SUBAPPLICATION SoftKeySR_PC_B_OPC_LOC (* Wie SoftKeySR_PC_B_OPC, aber Zustand lokal per PUBLISH (ein Geraet, Methoden per localhost) *)
  (* Standard: 61499-2; Description: Copyright (c) 2026 Meisterschulen am Ostbahnhof This program and the accompanying materials are made available under the terms of the Eclipse Public License 2.0 which is available at https://www.eclipse.org/legal/epl-2.0/ SPDX-License-Identifier: EPL-2.0 *)
  (* Version 1.3, 2026-11-25, Franz Höpfinger, Meisterschulen am Ostbahnhof, SERVER_0 -> MyLib::net::SERVER_0_QO (IND nur bei QO=TRUE, RSP intern). Ein gescheitertes RSP meldet IND mit QO=FALSE, direkt IND->RSP ergab eine Endlosschleife. *)
  (* Version 1.2, 2026-10-18, Franz Höpfinger, Meisterschulen am Ostbahnhof, Lokale Variante von SoftKeySR_PC_B_OPC: lokales PUBLISH statt Remote-WRITE (CLIENT) *)
  (* Version 1.1, 2026-09-09, Franz Höpfinger, Meisterschulen am Ostbahnhof, Fix: beide SERVER_0.RSP waren nie verdrahtet - blockierten je bis zu 4s den OPC-UA-Server-Thread (haelt open62541s globalen serviceMutex), verzoegerte dadurch JEDE OPC-UA-Statusmeldung projektweit. IND->RSP direkt verdrahtet. Siehe OPC_UA_VERNETZUNG.md Punkt 12. *)
  (* Version 1.0, 2026-09-03, Franz Höpfinger, Meisterschulen am Ostbahnhof, initial API and implementation and/or initial documentation *)
  PACKAGE MyLib::sys;
  IMPORT logiBUS::io::DQ::logiBUS_DO;
  IMPORT logiBUS::io::DQ::logiBUS_DO_S;
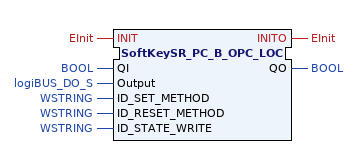
  EVENT_INPUT
    INIT : EInit; (* Initialization Request *)
  END_EVENT
  EVENT_OUTPUT
    INITO : EInit; (* Initialization Confirm *)
  END_EVENT
  VAR_INPUT
    QI : BOOL := TRUE; (* Quality Input - TRUE to enable service *)
    Output : logiBUS::io::DQ::logiBUS_DO_S := logiBUS_DO::Invalid; (* Identify the Output Output_Q1..Q8 *)
    ID_SET_METHOD : WSTRING; (* Lokale Methodenadresse (ACTION=CREATE_METHOD) fuer den Set-Methodenaufruf, wird von Geraet A per CALL_METHOD aufgerufen *)
    ID_RESET_METHOD : WSTRING; (* Lokale Methodenadresse (ACTION=CREATE_METHOD) fuer den Reset-Methodenaufruf, wird von Geraet A per CALL_METHOD aufgerufen *)
    ID_STATE_WRITE : WSTRING; (* Lokale Knotenadresse (BOOL, ACTION=WRITE) fuer den Zustand *)
  END_VAR
  VAR_OUTPUT
    QO : BOOL; (* Quality Output - TRUE if service executed successfully *)
  END_VAR
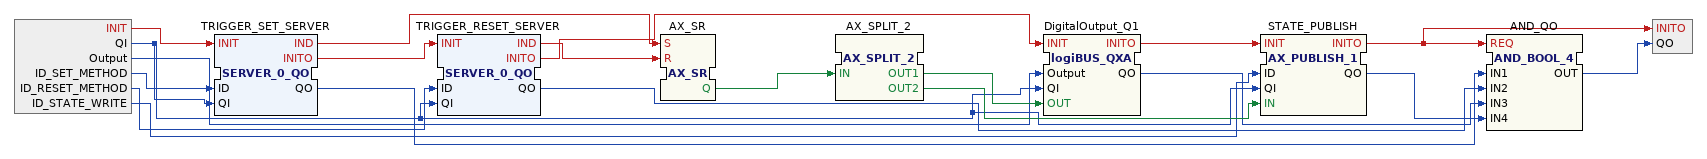
  FBS
    AX_SR : adapter::events::unidirectional::AX_SR;
    AX_SPLIT_2 : adapter::events::unidirectional::AX_SPLIT_2;
    DigitalOutput_Q1 : logiBUS::io::DQ::logiBUS_QXA;
    STATE_PUBLISH : adapter::net::AX_PUBLISH_1;
    AND_QO : iec61131::booleanOperators::AND_BOOL_4;
  END_FBS
  SUBAPPS
    TRIGGER_SET_SERVER : MyLib::net::SERVER_0_QO;
    TRIGGER_RESET_SERVER : MyLib::net::SERVER_0_QO;
  END_SUBAPPS
  EVENT_CONNECTIONS
    TRIGGER_SET_SERVER.IND TO AX_SR.S;
    TRIGGER_RESET_SERVER.IND TO AX_SR.R;
    INIT TO TRIGGER_SET_SERVER.INIT;
    TRIGGER_SET_SERVER.INITO TO TRIGGER_RESET_SERVER.INIT;
    TRIGGER_RESET_SERVER.INITO TO DigitalOutput_Q1.INIT;
    DigitalOutput_Q1.INITO TO STATE_PUBLISH.INIT;
    STATE_PUBLISH.INITO TO INITO;
    STATE_PUBLISH.INITO TO AND_QO.REQ;
  END_CONNECTIONS
  DATA_CONNECTIONS
    Output TO DigitalOutput_Q1.Output;
    ID_SET_METHOD TO TRIGGER_SET_SERVER.ID;
    ID_RESET_METHOD TO TRIGGER_RESET_SERVER.ID;
    ID_STATE_WRITE TO STATE_PUBLISH.ID;
    QI TO TRIGGER_SET_SERVER.QI;
    QI TO TRIGGER_RESET_SERVER.QI;
    QI TO DigitalOutput_Q1.QI;
    QI TO STATE_PUBLISH.QI;
    TRIGGER_SET_SERVER.QO TO AND_QO.IN1;
    TRIGGER_RESET_SERVER.QO TO AND_QO.IN2;
    DigitalOutput_Q1.QO TO AND_QO.IN3;
    STATE_PUBLISH.QO TO AND_QO.IN4;
    AND_QO.OUT TO QO;
  END_CONNECTIONS
  ADAPTER_CONNECTIONS
    AX_SR.Q TO AX_SPLIT_2.IN;
    AX_SPLIT_2.OUT1 TO DigitalOutput_Q1.OUT;
    AX_SPLIT_2.OUT2 TO STATE_PUBLISH.IN;
  END_CONNECTIONS
END_SUBAPPLICATION
